TYPE ST_VFDFunctions :
STRUCT
	Enable		: FB_SequencerFunction;
	LatchJogFwd : FB_SequencerFunction;
	LatchJogRev : FB_SequencerFunction;
	Stop 		: FB_SequencerFunction;
END_STRUCT
END_TYPE

(* stored: Version 1.1.0.1, ProductVersion 3.1.4024.12
   DUT ST_VFDFunctions: Id {b7685f85-c43b-4dc8-89e4-3fca04a5485c} *)
